Fanuc KAREL source: KC00008.KL

PROGRAM KC00008
%NOLOCKGROUP
%ENVIRONMENT PATHOP
VAR
  I: INTEGER
  J: INTEGER
  K: INTEGER
  R: REAL
  B: BOOLEAN
  S: STRING[80]
  T: STRING[80]
  P: PATH
  Q: PATH
  AI: ARRAY[8] OF INTEGER
  AB: ARRAY[244] OF BYTE
BEGIN
  DELETE_NODE(P,I,J)
END KC00008
